(* IEC 61131-3 sources: repolevel_ST_code_completion/output/0122完整版本_无planner目前sota/repoeval_open-type_dual-axis_winding_machine/readful_result_no_provide, 5 files *)

(* ---- CheckF.st ---- *)
VAR
END_VAR

IF lH <> 0 THEN
    lF := 9.8 * lM / (2 * COS(ATAN(lL / lH)));
ELSE
    lF := 0;
END_IF;
END_FUNCTION_BLOCK

(* ---- F_CalculateRadius.st ---- *)
F_CalculateRadius := ABS(SQRT(EXPT(lD, 2) + EXPT(lHnew + lOffset, 2)) - SQRT(EXPT(lD, 2) + EXPT(lHold + lOffset, 2))) / SMC_PI + lTk;
RETURN;
END_FUNCTION

(* ---- F_CompensateVelocity.st ---- *)
VAR
    lDeltaPos : LREAL; // Position change
END_VAR

// Calculate position change
lDeltaPos := lNewPos - lOldPos;

// Check if the axis is moving (position change)
IF lDeltaPos <> 0 THEN
    IF bUnwinding THEN
        // Unwinding: radius decreases, velocity needs to increase
        // Formula: V_new = V_old + V_old * Tk / (R - Tk)
        IF (lRadius - lTk) > 0.01 THEN // Avoid division by zero
            F_CompensateVelocity := lCurrentVel + lCurrentVel * lTk / (lRadius - lTk);
        ELSE
            F_CompensateVelocity := lCurrentVel;
        END_IF
    ELSE
        // Rewinding: radius increases, velocity needs to decrease
        // Formula: V_new = V_old - V_old * Tk / (R + Tk)
        IF (lRadius + lTk) > 0.01 THEN // Avoid division by zero
            F_CompensateVelocity := lCurrentVel - lCurrentVel * lTk / (lRadius + lTk);
        ELSE
            F_CompensateVelocity := lCurrentVel;
        END_IF
    END_IF
ELSE
    // Position unchanged, maintain current velocity
    F_CompensateVelocity := lCurrentVel;
END_IF;

RETURN;
END_FUNCTION

(* ---- SeekHome.st ---- *)
VAR
	_fbMoveVel	:	MC_MoveVelocity;
	_fbMoveAbs	:	MC_MoveAbsolute;
	_fbHalt		:	MC_Halt;
	_fbSetPos	:	MC_SetPosition;
	_fbRtrig	:	R_TRIG;
	_fbFtrig	:	F_TRIG;
	_nBDirection	:	MC_DIRECTION;
	_fTempPos		:	LREAL;
	_nState		:	USINT;
	_xPrevHome	:	BOOL;
	_xPrevAbort	:	BOOL;
	_xRefSwitchPrev	:	BOOL;
	_xIndexPulsePrev	:	BOOL;
END_VAR

IF _xAbort THEN
	_fbHalt.Execute := TRUE;
	_fbHalt.Axis := _Axis;
	_xBusy := FALSE;
	_xDone := FALSE;
	_xErr := FALSE;
	_iErrId := 0;
	_nState := 0;
	RETURN;
END_IF

CASE _nState OF
	0: // Idle
		IF _xHome THEN
			_xBusy := TRUE;
			_xDone := FALSE;
			_xErr := FALSE;
			_iErrId := 0;
			_nState := 1;
		END_IF;

	1: // Start Homing
		_fbMoveVel.Execute := TRUE;
		_fbMoveVel.Axis := _Axis;
		_fbMoveVel.Velocity := _fFastHomeVel;
		_fbMoveVel.Acceleration := _fHomeAcc;
		_fbMoveVel.Deceleration := _fHomeDec;
		_fbMoveVel.Direction := _nDirection;

		IF _xReferenceSwitch THEN
			_fbMoveVel.Execute := FALSE;
			_nState := 2;
		END_IF;

	2: // Slow Homing
		_fbMoveVel.Execute := TRUE;
		_fbMoveVel.Velocity := _fSlowHomeVel;

		IF _xIndexPulse THEN
			_fbMoveVel.Execute := FALSE;
			_nState := 3;
		END_IF;

	3: // Set Position
		_fbSetPos.Execute := TRUE;
		_fbSetPos.Axis := _Axis;
		_fbSetPos.Position := _fHomePos;

		IF NOT _fbSetPos.Busy THEN
			_fbSetPos.Execute := FALSE;
			_xBusy := FALSE;
			_xDone := TRUE;
			_nState := 0;
		END_IF;

	ELSE
		_xErr := TRUE;
		_iErrId := 1; // Error code for unexpected state
		_xBusy := FALSE;
		_nState := 0;
	END_CASE;
RETURN;
END_FUNCTION_BLOCK

(* ---- StaDisplay.st ---- *)
VAR
END_VAR

CASE iStatus OF
	2,3,4,5,6,7,8,9,10,221,222:
		Y5 := FALSE;
		Y6 := TRUE;
		Y1 := TRUE;
		Y2 := FALSE;
		Y3 := FALSE;
		Y4 := FALSE;
	11,12:
		Y5 := FALSE;
		Y6 := TRUE;
		Y1 := FALSE;
		Y2 := TRUE;
		Y3 := FALSE;
		Y4 := FALSE;
	13,14,15,16,17,18,19,20,21,22:
		Y5 := TRUE;
		Y6 := FALSE;
		Y1 := FALSE;
		Y2 := FALSE;
		Y3 := TRUE;
		Y4 := FALSE;
	23,24:
		Y5 := TRUE;
		Y6 := FALSE;
		Y1 := FALSE;
		Y2 := FALSE;
		Y3 := FALSE;
		Y4 := TRUE;
	ELSE
		Y5 := FALSE;
		Y6 := FALSE;
		Y1 := FALSE;
		Y2 := FALSE;
		Y3 := FALSE;
		Y4 := FALSE;
END_CASE;
END_FUNCTION_BLOCK
